Staubli VAL3: start.pgx

public program start()
begin
  if prog:libLoad("./LongProg")!=0
    logMsg("Error Loading RoboDK library")
    popUpMsg("Error Loading RoboDK library")
  endIf
  wait(taskStatus("loading")==-1)
  taskCreate "loading",10,loadNextOne("./LongProg2")
  call prog:start()

  if prog:libLoad("./LongProg2")!=0
    logMsg("Error Loading RoboDK library")
    popUpMsg("Error Loading RoboDK library")
  endIf
  wait(taskStatus("loading")==-1)
  taskCreate "loading",10,loadNextOne("./LongProg3")
  call prog:start()

  if prog:libLoad("./LongProg3")!=0
    logMsg("Error Loading RoboDK library")
    popUpMsg("Error Loading RoboDK library")
  endIf
  wait(taskStatus("loading")==-1)
  call prog:start()


end
